                   IF NOT #found THEN
                       #VarErr := 1;                       // no feasible transfer
                   ELSIF #CurLen >= 96 THEN
                       #VarErr := 2;                       // plan longer than 96 transfers
                   ELSE
                       // ---------- apply the best (s, d) ----------
                       #si := #bS;
                       #sCol := #SrcX[#si];
                       #sRow := #SrcY[#si];
                       #sBay := #SrcB[#si];
                       #dBay := #bDb;
                       #dCol := #FreeX[#dBay, #bK];
                       #dRow := #FreeY[#dBay, #bK];
                       #eT := "Crane_MoveCost"(X0 := #cx, Y0 := #cy, B0 := #cb, X1 := #sCol, Y1 := #sRow, B1 := #sBay,
                                               MMode := #cMMode, M => #eMan);
                       #lT := "Crane_MoveCost"(X0 := #sCol, Y0 := #sRow, B0 := #sBay, X1 := #dCol, Y1 := #dRow, B1 := #dBay,
                                               MMode := #cMMode, M => #lMan);
                       #g[#dBay, #dCol, #dRow] := #g[#sBay, #sCol, #sRow];
                       #g[#sBay, #sCol, #sRow] := 0;
                       #TotT := #TotT + #eT + 200 + #lT + 200;
                       #TotM := #TotM + INT_TO_DINT(#eMan) + 1 + INT_TO_DINT(#lMan) + 1;
                       #CurLen := #CurLen + 1;
                       #CurPlan[#CurLen].Kind := #SrcKind[#si];
                       #CurPlan[#CurLen].Id := #SrcId[#si];
                       #CurPlan[#CurLen].ListIdx := #SrcIdx[#si];
                       #CurPlan[#CurLen].SrcX := INT_TO_SINT(#sCol);
                       #CurPlan[#CurLen].SrcY := INT_TO_SINT(#sRow);
                       #CurPlan[#CurLen].SrcBay := INT_TO_USINT(#sBay);
                       #CurPlan[#CurLen].DstX := INT_TO_SINT(#dCol);
                       #CurPlan[#CurLen].DstY := INT_TO_SINT(#dRow);
                       #CurPlan[#CurLen].DstBay := INT_TO_USINT(#dBay);
                       #CurPlan[#CurLen].CumT_ds := #TotT;
                       #CurPlan[#CurLen].CumM := #TotM;
                       #CurSrc[#CurLen] := #si;
                       #cx := #dCol;
                       #cy := #dRow;
                       #cb := #dBay;
                       #cG := #FreeG[#dBay, #bK];
                       #Pend[#si] := FALSE;
                       #nPend := #nPend - 1;
                   END_IF;
               END_IF;

               IF #PubPending THEN
                   // ---------- job finished: publish (World is written only here) ----------
                   #PubPending := FALSE;
                   IF #HaveBest THEN
                       FOR #i := 1 TO 96 DO
                           IF #i <= #BestLen THEN
                               "World".Plan[#i] := #BestPlan[#i];
                           ELSE
                               "World".Plan[#i] := #ZeroTr;
                           END_IF;
                       END_FOR;
                       "World".PlanLen := #BestLen;
                       "World".PlanVariant := #BestV;
                       "World".PredT_ds := #BestT;
                       "World".PredM := #BestM;
                       "World".LbT_ds := #sBaseT + #LbT;
                       "World".LbM := #sBaseM + #LbM;
                       "World".ImpEvals := #ImpEvals;
                       "World".ImpAccepts := #ImpAcc;
                       "World".SlotAccepts := #SlAcc;
                       "World".OrderFeasible := #OrderOk;
                       IF #sN > 0 THEN
                           "World".PredJ := 0.5 * (DINT_TO_REAL(#BestT) / 10.0) / (76.0 * INT_TO_REAL(#sN))
                                          + 0.5 * DINT_TO_REAL(#BestM) / (4.0 * INT_TO_REAL(#sN));
                           "World".PredJ0 := 0.5 * (DINT_TO_REAL(#GrT) / 10.0) / (76.0 * INT_TO_REAL(#sN))
                                           + 0.5 * DINT_TO_REAL(#GrM) / (4.0 * INT_TO_REAL(#sN));
                           "World".LbJ := 0.5 * (DINT_TO_REAL(#sBaseT + #LbT) / 10.0) / (76.0 * INT_TO_REAL(#sN))
                                        + 0.5 * DINT_TO_REAL(#sBaseM + #LbM) / (4.0 * INT_TO_REAL(#sN));
                       ELSE
                           "World".PredJ := 0.0;
                           "World".PredJ0 := 0.0;
                           "World".LbJ := 0.0;
                       END_IF;
                       "World".PlanValid := TRUE;
                       #Done := TRUE;
                       #ErrCode := 0;
                   ELSE
                       "World".PlanValid := FALSE;
                       "World".PlanLen := 0;
                       "World".PlanVariant := 0;
                       "World".SlotAccepts := 0;
                       "World".OrderFeasible := #OrderOk;
                       #Error := TRUE;
                       #ErrCode := #Err1;
                   END_IF;
                   #JobBusy := FALSE;
               END_IF;
           END_WHILE;
           #DiagCallMs := RUNTIME(MEM := #RtMem) * 1000.0;
           #DiagJobMs := #DiagJobMs + #DiagCallMs;
           IF #DiagCallMs > #DiagMaxCallMs THEN
               #DiagMaxCallMs := #DiagCallMs;
           END_IF;
       END_IF;
   END_REGION

   #Busy := #JobBusy;
END_FUNCTION_BLOCK

FUNCTION "CheckCmd" : Int   // FC10, SCL
TITLE = Pre-check of a crane command before OB30 issues it to FB1
{ S7_Optimized_Access := 'TRUE' }
VERSION : 0.1
// Returns 0 = OK, otherwise the alarm bit number (CONTRACT 1.4 / 3.3):
//     100 ship imbalance (alarm bit 0)      1 pick location empty
//       2 drop location occupied            9 invalid command / position
//      11 crane already carrying (lift, or MANUAL reset with a load)   12 crane is empty (put down)
//   The first failing rule decides the result.
//   Lift/put act on the CURRENT crane position (CraneX/Y/Bay); the X/Y/Bay of C are ignored.
//   Balance rule (CONTRACT 4.3 step rule): the result is OK if |L'-R'| <= BalLimit,
//   or if it is not worse than before (|L'-R'| <= |L-R|). Same for front/aft if BalMode = 1.
//   v1.5 (R2-J1): relaxed rule while "World".BalCeil > BalLimit (set by FB10 only when the ship started out
//   of balance and the list order is infeasible otherwise): while |L-R| > BalLimit, |L'-R'| <= BalCeil is OK.
   VAR_INPUT
      C : "typeCmd";   // command to check
      CraneX : SInt;   // crane position now
      CraneY : SInt;
      CraneBay : USInt;
      Carried : UInt;   // ID on the hook (0 = none)
      BalLimit : Int;   // max |L-R| (5)
      BalMode : USInt;   // 0 left/right only, 1 also front/aft
   END_VAR
   VAR_TEMP
      x : Int;
      y : Int;
      cx : Int;
      cy : Int;
      cell : UInt;
      delta : Int;   // -1 lift (container leaves the ship), +1 put
      L : Int;   // ship count x in {0,1}
      R : Int;   // ship count x in {2,3}
      F : Int;   // ship count y in 0..5
      "A" : Int;   // ship count y in 6..11
      L2 : Int;
      R2 : Int;
      F2 : Int;
      A2 : Int;
   END_VAR
BEGIN
   REGION Move and reset
       CASE #C.Cmd OF
           3:  // move to (X, Y, Bay): only the target must be a valid slot
               IF #C.X >= 0 AND #C.X <= 3 AND #C.Y >= 0 AND #C.Y <= 11 AND #C.Bay <= 1 THEN
                   #CheckCmd := 0;
               ELSE
                   #CheckCmd := 9;
               END_IF;
               RETURN;
           10: // reset of FB1: INIT may always reset (it reloads the yard and clears the hook);
               // a MANUAL reset with a container on the hook would lose it and the score counters
               IF #C.Src = 3 AND #Carried <> 0 THEN
                   #CheckCmd := 11;
               ELSE
                   #CheckCmd := 0;
               END_IF;
               RETURN;
           1, 2:
               ;   // checked below
           ELSE
               #CheckCmd := 9;
               RETURN;
       END_CASE;
   END_REGION

   REGION Lift / put: crane position and hook
       #cx := SINT_TO_INT(#CraneX);
       #cy := SINT_TO_INT(#CraneY);
       IF #cx < 0 OR #cx > 3 OR #cy < 0 OR #cy > 11 OR #CraneBay > 1 THEN
           #CheckCmd := 9;     // crane is not over a valid slot
           RETURN;
       END_IF;

       IF #CraneBay = 0 THEN
           #cell := "World".Bay0[#cx, #cy];
       ELSE
           #cell := "World".Bay1[#cx, #cy];
       END_IF;

       IF #C.Cmd = 1 THEN
           IF #Carried <> 0 THEN
               #CheckCmd := 11;    // already carrying a container
               RETURN;
           END_IF;
           IF #cell = 0 THEN
               #CheckCmd := 1;     // pick location empty
               RETURN;
           END_IF;
           #delta := -1;
       ELSE
           IF #Carried = 0 THEN
               #CheckCmd := 12;    // nothing on the hook
               RETURN;
           END_IF;
           IF #cell <> 0 THEN
               #CheckCmd := 2;     // drop location occupied
               RETURN;
           END_IF;
           #delta := 1;
       END_IF;
   END_REGION

   REGION Ship balance after the lift / put (only when it happens on the ship)
       IF #CraneBay = 0 THEN
           #L := 0; #R := 0; #F := 0; #A := 0;
           FOR #x := 0 TO 3 DO
               FOR #y := 0 TO 11 DO
                   IF "World".Bay0[#x, #y] <> 0 THEN
                       IF #x <= 1 THEN #L := #L + 1; ELSE #R := #R + 1; END_IF;
                       IF #y <= 5 THEN #F := #F + 1; ELSE #A := #A + 1; END_IF;
                   END_IF;
               END_FOR;
           END_FOR;

           #L2 := #L; #R2 := #R; #F2 := #F; #A2 := #A;
           IF #cx <= 1 THEN #L2 := #L + #delta; ELSE #R2 := #R + #delta; END_IF;
           IF #cy <= 5 THEN #F2 := #F + #delta; ELSE #A2 := #A + #delta; END_IF;

           IF ABS(#L2 - #R2) > #BalLimit AND ABS(#L2 - #R2) > ABS(#L - #R)
               AND NOT (ABS(#L - #R) > #BalLimit AND ABS(#L2 - #R2) <= "World".BalCeil)
           THEN
               #CheckCmd := 100;
               RETURN;
           END_IF;
           IF #BalMode = 1 AND ABS(#F2 - #A2) > #BalLimit AND ABS(#F2 - #A2) > ABS(#F - #A) THEN
               #CheckCmd := 100;
               RETURN;
           END_IF;
       END_IF;

       #CheckCmd := 0;
   END_REGION
END_FUNCTION

FUNCTION "Crane_MoveCost" : DInt   // FC20, SCL
TITLE = Time and manipulation cost of one crane move (CONTRACT 4.1)
{ S7_Optimized_Access := 'TRUE' }
VERSION : 0.1
// Returns the move time in DECISECONDS (DInt) from (X0,Y0,B0) to (X1,Y1,B1); output M = manipulations.
//   Global column G(x, b) = x + 6 for bay 0 (ship), x for bay 1 (yard)   (one yard bay only).
//   Same position              -> T = 0, M = 0
//   otherwise                  -> T = max(60*|dG|, 23*|dy|) ds   (6 m per column / 2.3 m per row at 1 m/s)
//   MMode 0 (spec, global X)   -> M = [dG <> 0] + [dy <> 0]
//   MMode 1 (local x)          -> M = [x1 <> x0] + [dy <> 0]
//   MMode 2 (per command, FB1) -> M = 1
//   Any other MMode is treated as 0. No range checks: callers pass valid positions
//   (the planner also uses it with synthetic columns 0..9 in bay 1 to build its cost table).
   VAR_INPUT
      X0 : Int;
      Y0 : Int;
      B0 : Int;
      X1 : Int;
      Y1 : Int;
      B1 : Int;
      MMode : Int;
   END_VAR
   VAR_OUTPUT
      "M" : Int;
   END_VAR
   VAR_TEMP
      g0 : DInt;
      g1 : DInt;
      dG : DInt;
      dY : DInt;
      tX : DInt;
      tY : DInt;
   END_VAR
BEGIN

    // Zero move: no time, no manipulation (the runtime never issues it, U6).
    IF #X0 = #X1 AND #Y0 = #Y1 AND #B0 = #B1 THEN
        #M := 0;
        #Crane_MoveCost := 0;
        RETURN;
    END_IF;

    // Global columns
    #g0 := INT_TO_DINT(#X0);
    IF #B0 = 0 THEN
        #g0 := #g0 + 6;
    END_IF;
    #g1 := INT_TO_DINT(#X1);
    IF #B1 = 0 THEN
        #g1 := #g1 + 6;
    END_IF;
    #dG := ABS(#g1 - #g0);
    #dY := ABS(INT_TO_DINT(#Y1) - INT_TO_DINT(#Y0));

    // Time: both axes travel at the same time, the longer one decides
    #tX := 60 * #dG;
    #tY := 23 * #dY;
    IF #tX >= #tY THEN
        #Crane_MoveCost := #tX;
    ELSE
        #Crane_MoveCost := #tY;
    END_IF;

    // Manipulations
    #M := 0;
    CASE #MMode OF
        1:
            IF #X1 <> #X0 THEN
                #M := #M + 1;
            END_IF;
            IF #dY <> 0 THEN
                #M := #M + 1;
            END_IF;
        2:
            #M := 1;
        ELSE
            IF #dG <> 0 THEN
                #M := #M + 1;
            END_IF;
            IF #dY <> 0 THEN
                #M := #M + 1;
            END_IF;
    END_CASE;
END_FUNCTION

FUNCTION "Crane_DropCost" : DInt   // FC21, SCL
TITLE = Weighted cost of a drop cell in the planner SLOT phase (CONTRACT 4.11)
{ S7_Optimized_Access := 'TRUE' }
VERSION : 0.1
// c(d) = W(source -> cell) + W(cell -> next source)   (second term only if HasNxt)
//   W = T [ds] + 190 * M, both from FC20 "Crane_MoveCost" (the only cost formula).
//   Python reference: tools/crane_plan.py slot_search() cost(); mirror tia-src/13_improve_mirror.py.
   VAR_INPUT
      SrcX : Int;
      SrcY : Int;
      SrcB : Int;
      CelX : Int;
      CelY : Int;
      CelB : Int;
      NxtX : Int;
      NxtY : Int;
      NxtB : Int;
      HasNxt : Bool;
      MMode : Int;
   END_VAR
   VAR_TEMP
      tA : DInt;
      mA : Int;
      wSum : DInt;
   END_VAR
BEGIN

    #tA := "Crane_MoveCost"(X0 := #SrcX, Y0 := #SrcY, B0 := #SrcB, X1 := #CelX, Y1 := #CelY, B1 := #CelB,
                            MMode := #MMode, M => #mA);
    #wSum := #tA + 190 * INT_TO_DINT(#mA);
    IF #HasNxt THEN
        #tA := "Crane_MoveCost"(X0 := #CelX, Y0 := #CelY, B0 := #CelB, X1 := #NxtX, Y1 := #NxtY, B1 := #NxtB,
                                MMode := #MMode, M => #mA);
        #wSum := #wSum + #tA + 190 * INT_TO_DINT(#mA);
    END_IF;
    #Crane_DropCost := #wSum;
END_FUNCTION

ORGANIZATION_BLOCK "Main"   // OB1, SCL, ProgramCycle
TITLE = "Main Program Sweep (Cycle)"
{ S7_Optimized_Access := 'TRUE' }
VERSION : 0.1
   VAR_INPUT
      Initial_Call : Bool;   // Initial call of this OB
      Remanence : Bool;   // =True, if remanent data are available
   END_VAR
BEGIN

    // Crane control (FB10): modes, state machine, planning, HMI interface.
    // FB1 "Crane_manipulation" is called only in OB30 "Cyclic interrupt" (1 s).
    "Crane_Control_DB"();
END_ORGANIZATION_BLOCK

ORGANIZATION_BLOCK "Cyclic interrupt"   // OB30, SCL, CyclicInterrupt
TITLE = Crane command execution (1 s cyclic interrupt)
{ S7_Optimized_Access := 'TRUE' }
VERSION : 0.1
   VAR_INPUT
      Initial_Call : Bool;   // Initial call of this OB
      Event_Count : Int;   // Events discarded
   END_VAR
   VAR_TEMP
      rc : Int;   // result of "CheckCmd"
      bitNo : Int;   // alarm bit to set in "World".Fault
      cx : Int;
      cy : Int;
      gxOld : Int;   // global column before / after a move (Bay0 x + 6, Bay1 x)
      gxNew : Int;
      cmd : "typeCmd";   // command to issue
   END_VAR
BEGIN
   // OB30 runs every 1 s (spec: "once per second"). It is the ONLY place that
   // calls FB1 "Crane_manipulation" and writes its command tags MB100..MB103.
   // FB10 "Crane_Control" (OB1) decides WHAT to do and stages it in "World".NextCmd;
   // OB30 decides WHEN: only after FB1 reported the previous command finished
   // (command_id back to 0) and only after "CheckCmd" accepted the command.
   // Order per tick (CONTRACT 3.4): 1 tick, 2 completion, 3 issue, 4 FB1 call.

   REGION 1 Tick counter and heartbeat
       "World".OB30Ticks := "World".OB30Ticks + 1;
       "HMI_IF".Heartbeat := NOT "HMI_IF".Heartbeat;
   END_REGION

   REGION 2 Has the previous command finished?
       IF "World".Busy THEN
           IF "new_command_ID" = 0 THEN
               // Spec section 3 manipulation count (shown next to FB1's MD107):
               // a move counts +1 per changed axis (x incl. bay change, y), lift / put +1, reset clears
               CASE "World".ActCmd.Cmd OF
                   1, 2:
                       "World".MSpec := "World".MSpec + 1;
                   3:
                       #gxOld := SINT_TO_INT("World".CraneX);
                       IF "World".CraneBay = 0 THEN #gxOld := #gxOld + 6; END_IF;
                       #gxNew := SINT_TO_INT("x_position");
                       IF "bay_ID" = 0 THEN #gxNew := #gxNew + 6; END_IF;
                       IF #gxNew <> #gxOld THEN "World".MSpec := "World".MSpec + 1; END_IF;
                       IF "y_position" <> "World".CraneY THEN "World".MSpec := "World".MSpec + 1; END_IF;
                   10:
                       "World".MSpec := 0;
                   ELSE
                       ;
               END_CASE;

               // FB1 finished: take over the crane position it reports
               "World".CraneX := "x_position";
               "World".CraneY := "y_position";
               "World".CraneBay := "bay_ID";

               // Effect of the command on our container model (FB1 does not track containers)
               #cx := SINT_TO_INT("World".ActCmd.X);
               #cy := SINT_TO_INT("World".ActCmd.Y);
               CASE "World".ActCmd.Cmd OF
                   1:  // lift: the container moves from the cell to the hook
                       IF #cx >= 0 AND #cx <= 3 AND #cy >= 0 AND #cy <= 11 THEN
                           IF "World".ActCmd.Bay = 0 THEN
                               "World".Carried := "World".Bay0[#cx, #cy];
                               "World".Bay0[#cx, #cy] := 0;
                           ELSIF "World".ActCmd.Bay = 1 THEN
                               "World".Carried := "World".Bay1[#cx, #cy];
                               "World".Bay1[#cx, #cy] := 0;
                           END_IF;
                       END_IF;
                   2:  // put down: the container moves from the hook to the cell
                       IF #cx >= 0 AND #cx <= 3 AND #cy >= 0 AND #cy <= 11 THEN
                           IF "World".ActCmd.Bay = 0 THEN
                               "World".Bay0[#cx, #cy] := "World".Carried;
                               "World".Carried := 0;
                           ELSIF "World".ActCmd.Bay = 1 THEN
                               "World".Bay1[#cx, #cy] := "World".Carried;
                               "World".Carried := 0;
                           END_IF;
                       END_IF;
                   3:  // move: FB1 must now report the commanded position
                       IF "World".CraneX <> "World".ActCmd.X
                           OR "World".CraneY <> "World".ActCmd.Y
                           OR "World".CraneBay <> "World".ActCmd.Bay
                       THEN
                           "World".Fault := "World".Fault OR WORD#16#4000;   // bit 14 position mismatch
                       END_IF;
                   ELSE
                       ;   // 10 reset: the crane position comes from FB1 (0,0,1)
               END_CASE;

               "World".LastDone := "World".ActCmd;
               "World".DoneSeq := "World".DoneSeq + 1;
               "World".Busy := FALSE;
               "World".BusyTicks := 0;
           ELSE
               // Still executing: watchdog
               IF "World".BusyTicks < 32000 THEN
                   "World".BusyTicks := "World".BusyTicks + 1;
               END_IF;
               IF "World".BusyTicks > "World".CfgTimeoutTicks THEN
                   "World".Fault := "World".Fault OR WORD#16#0400;           // bit 10 FB1 timeout
               END_IF;
           END_IF;
       END_IF;
   END_REGION

   REGION 3 Issue the next command (only when the previous one is done)
       // Spec 2.2: "na pocetku bloka OB30 provjeriti je li posljednja manipulacija izvrsena":
       // FB1 resets "new_command_ID" (MB103) to 0 when a command is done (checked in region 2
       // for World.Busy and here again literally, so a stray MB103 value is never overwritten).
       IF NOT "World".Busy AND "new_command_ID" = 0 AND "World".CmdReady AND "World".Permit AND "World".Fault = 0 THEN
           #cmd := "World".NextCmd;
           // Lift / put always act where the crane is now
           IF #cmd.Cmd = 1 OR #cmd.Cmd = 2 THEN
               #cmd.X := "World".CraneX;
               #cmd.Y := "World".CraneY;
               #cmd.Bay := "World".CraneBay;
           END_IF;

           // Pick not empty, drop not occupied, slot valid, ship stays balanced
           #rc := "CheckCmd"(C := #cmd,
                             CraneX := "World".CraneX,
                             CraneY := "World".CraneY,
                             CraneBay := "World".CraneBay,
                             Carried := "World".Carried,
                             BalLimit := "World".CfgBalLimit,
                             BalMode := "World".CfgBalMode);

           IF #rc = 0 THEN
               "new_x_position" := #cmd.X;
               "new_y_position" := #cmd.Y;
               "new_bay_ID" := #cmd.Bay;
               "new_command_ID" := #cmd.Cmd;
               "World".ActCmd := #cmd;
               "World".Busy := TRUE;
               "World".BusyTicks := 0;
           ELSE
               // Rejected: raise the alarm and do not issue (halts until ACK in FB10)
               IF #rc = 100 THEN
                   #bitNo := 0;
               ELSE
                   #bitNo := #rc;
               END_IF;
               IF #bitNo >= 0 AND #bitNo <= 15 THEN
                   "World".Fault := "World".Fault OR SHL(IN := WORD#16#0001, N := INT_TO_UINT(#bitNo));
               ELSE
                   "World".Fault := "World".Fault OR WORD#16#0200;           // unknown code -> bit 9
               END_IF;
               "World".FaultCmd := #cmd;
           END_IF;
           "World".CmdReady := FALSE;
       END_IF;
   END_REGION

   REGION 4 FB1 call (every tick; command 0 = nothing to do)
       "Crane_manipulation_DB"(new_x_position := "new_x_position",
                               new_y_position := "new_y_position",
                               new_bay_ID := "new_bay_ID",
                               pos_x_after_command => "x_position",
                               pos_y_after_command => "y_position",
                               bay_ID_after_command => "bay_ID",
                               number_of_manipulations => "number_of_manipulations",
                               working_time => "time",
                               command_id := "new_command_ID");
   END_REGION
END_ORGANIZATION_BLOCK

ORGANIZATION_BLOCK "Startup"   // OB100, SCL, Startup
TITLE = "Complete Restart"
{ S7_Optimized_Access := 'TRUE' }
VERSION : 0.1
   VAR_INPUT
      LostRetentive : Bool;   // True if retentive data are lost
      LostRTC : Bool;   // True if date and time are lost
   END_VAR
BEGIN
   // define the inital state of the shipyard
   "Crane_manipulation_DB".command_id := 0; // set "do nothing" command
   "Crane_manipulation_DB".current_bay_ID := 1; // the crane starting bay ID set to 1 (left of the ship)
   "Crane_manipulation_DB".current_x_position_in_bay := 0; // starting X position of the crane
   "Crane_manipulation_DB".current_y_position_in_bay := 0; // starting Y position of the crane

   //define startup command parameters
   "new_x_position" := 0; // starting X position of the crane
   "new_y_position" := 0; // starting Y position of the crane
   "new_bay_ID" := 1; // the crane starting bay ID set to 1 (left of the ship)
   "new_command_ID" := 0; // set "do nothing" command

   // reset of evaluation parameters
   "Crane_manipulation_DB".total_number_of_manipulations := 0; // reset total number of the crane manipulations
   "Crane_manipulation_DB".total_time := 0.0; // reset of total time
END_ORGANIZATION_BLOCK

(* ===== HMI "HMI_RT_1" =====
connection "HMI_Connection_1": ETHERNET, S7_1500_OMS

HMI tags "Default tag table"
   "time" : Real = PLC time AT %MD112, 1 s

screen "Screen_1" 1024x768
   TextField "Text field_1" at 20,17 size 95x22; Text 'PLC+ 2019:'
   IOField "I/O field_1" at 86,66 size 96x32; FormatPattern s999999999.999
      ProcessValue <- "time"
*)